(* IEC 61131-3 sources: test/Class/HmiScreen, 1 file *)

(* ---- HmiScreen.st ---- *)
#include "..\..\Source\Common\hmi_nuc.h"

(*!
<Class
	Name               = "HmiScreen"
	Revision           = "0.1"
	RealtimeTask       = "false"
	CyclicTask         = "false"
	BackgroundTask     = "false"
	Sigmatek           = "true"
	OSInterface        = "false"
	HighPriority       = "false"
	Automatic          = "false"
	UpdateMode         = "Prescan"
	SharedCommandTable = "true"
	Objectsize         = "(284,120)">
	<Channels>
		<Client Name="MemCircle" Required="true" Internal="true"/>
		<Client Name="MemImage" Required="true" Internal="true"/>
		<Client Name="MemIO" Required="true" Internal="true"/>
		<Client Name="MemLine" Required="true" Internal="true"/>
		<Client Name="MemRectangle" Required="true" Internal="true"/>
		<Client Name="MemText" Required="true" Internal="true"/>
		<Client Name="MemZorder" Required="true" Internal="true"/>
	</Channels>
	<Dependencies>
		<Files>
			<File Path=".\Source\Common\hmi_nuc.h" Include="true"/>
		</Files>
	</Dependencies>
	<RevDoku>
		<Owner Company="sigmatek" Author="kolott"/>
		<Dokumentation Revision="0.1" Date="2014-04-15" Author="kolott" Company="sigmatek" Description="new method FreeMem()"/>
	</RevDoku>
	<Network Name="HmiScreen">
		<!-- List of Components in this network -->
		<Components>
			<Object
				Name       = "_base"
				Class      = "HmiBaseList"
				Position   = "(218,120)"
				Visualized = "false">
				<Channels>
					<Server Name="ClassSvr"/>
					<Client Name="File"/>
				</Channels>
			</Object>
			<Object
				Name       = "MemCircle"
				Class      = "HmiMemCircle"
				Position   = "(600,510)"
				Visualized = "false">
				<Channels>
					<Server Name="ClassSvr"/>
					<Client Name="File"/>
				</Channels>
			</Object>
			<Object
				Name       = "MemImage"
				Class      = "HmiMemImage"
				Position   = "(600,810)"
				Visualized = "false">
				<Channels>
					<Server Name="ClassSvr"/>
					<Client Name="File"/>
				</Channels>
			</Object>
			<Object
				Name       = "MemIO"
				Class      = "HmiMemIO"
				Position   = "(210,810)"
				Visualized = "false">
				<Channels>
					<Server Name="ClassSvr"/>
					<Client Name="File"/>
				</Channels>
			</Object>
			<Object
				Name       = "MemLine"
				Class      = "HmiMemLine"
				Position   = "(600,660)"
				Visualized = "false">
				<Channels>
					<Server Name="ClassSvr"/>
					<Client Name="File"/>
				</Channels>
			</Object>
			<Object
				Name       = "MemRectangle"
				Class      = "HmiMemRectangle"
				Position   = "(210,510)"
				Visualized = "false">
				<Channels>
					<Server Name="ClassSvr"/>
					<Client Name="File"/>
				</Channels>
			</Object>
			<Object
				Name       = "MemText"
				Class      = "HmiMemText"
				Position   = "(210,660)"
				Visualized = "false">
				<Channels>
					<Server Name="ClassSvr"/>
					<Client Name="File"/>
				</Channels>
			</Object>
			<Object
				Name       = "MemZorder"
				Class      = "HmiMemZorder"
				Position   = "(450,330)"
				Visualized = "false">
				<Channels>
					<Server Name="ClassSvr"/>
					<Client Name="File"/>
				</Channels>
			</Object>
		</Components>
		<Comments>
		</Comments>
		<!-- List of Connections in this network -->
		<Connections>
			<Connection Source="this.ClassSvr" Destination="_base.ClassSvr" Vertices="(1072,210),(518,210),"/>
			<Connection Source="_base.File" Destination="this.File" Vertices="(218,210),(38,210),"/>
			<Connection Source="this.MemZorder" Destination="MemZorder.ClassSvr"/>
			<Connection Source="MemZorder.File" Destination="this.File" Vertices="(450,420),(38,210),"/>
			<Connection Source="this.MemRectangle" Destination="MemRectangle.ClassSvr"/>
			<Connection Source="MemRectangle.File" Destination="this.File" Vertices="(210,600),(38,210),"/>
			<Connection Source="this.MemText" Destination="MemText.ClassSvr"/>
			<Connection Source="MemText.File" Destination="this.File" Vertices="(210,750),(38,210),"/>
			<Connection Source="this.MemIO" Destination="MemIO.ClassSvr"/>
			<Connection Source="MemIO.File" Destination="this.File" Vertices="(210,900),(38,210),"/>
			<Connection Source="this.MemCircle" Destination="MemCircle.ClassSvr"/>
			<Connection Source="MemCircle.File" Destination="this.File" Vertices="(600,600),(38,210),"/>
			<Connection Source="this.MemLine" Destination="MemLine.ClassSvr"/>
			<Connection Source="MemLine.File" Destination="this.File" Vertices="(600,750),(38,210),"/>
			<Connection Source="this.MemImage" Destination="MemImage.ClassSvr"/>
			<Connection Source="MemImage.File" Destination="this.File" Vertices="(600,900),(38,210),"/>
		</Connections>
		<!-- Headerfiles -->
		<Options>
		</Options>
	</Network>
</Class>
*)
#pragma using HmiBaseList

HmiScreen : CLASS
: HmiBaseList
  //Servers:
  //Clients:
	MemRectangle 	: CltChCmd_HmiMemRectangle;
	MemText 	: CltChCmd_HmiMemText;
	MemIO 	: CltChCmd_HmiMemIO;
	MemCircle 	: CltChCmd_HmiMemCircle;
	MemLine 	: CltChCmd_HmiMemLine;
	MemImage 	: CltChCmd_HmiMemImage;
	MemZorder 	: CltChCmd_HmiMemZorder;
  //Variables:
		StartFunct 	: UDINT;
		EndFunct 	: UDINT;
  //Functions:

	FUNCTION VIRTUAL Load
		VAR_OUTPUT
			retcode 	: BOOL;
		END_VAR;

	FUNCTION VIRTUAL Free;

	FUNCTION GLOBAL GetZorder
		VAR_INPUT
			index 	: UDINT;
		END_VAR
		VAR_OUTPUT
			retcode 	: ^HMI_ANYTHING;
		END_VAR;

	FUNCTION GLOBAL GetZorderNo
		VAR_OUTPUT
			retcode 	: UDINT;
		END_VAR;

	FUNCTION GLOBAL GetControl
		VAR_INPUT
			pany 	: ^HMI_ANYTHING;
		END_VAR
		VAR_OUTPUT
			retcode 	: ^void;
		END_VAR;

	FUNCTION GLOBAL GetStartFunct
		VAR_OUTPUT
			retcode 	: UDINT;
		END_VAR;

	FUNCTION GLOBAL GetEndFunct
		VAR_OUTPUT
			retcode 	: UDINT;
		END_VAR;

	FUNCTION GLOBAL FreeMem;
  //Tables:
	FUNCTION @STD
		VAR_OUTPUT
			ret_code	: CONFSTATES;
		END_VAR;
	FUNCTION GLOBAL TAB @CT_;
END_CLASS;

#pragma using HmiMemCircle
#pragma using HmiMemImage
#pragma using HmiMemIO
#pragma using HmiMemLine
#pragma using HmiMemRectangle
#pragma using HmiMemText
#pragma using HmiMemZorder

FUNCTION VIRTUAL HmiScreen::Free

  MemZorder.Free();
  MemRectangle.Free();
  MemText.Free();
  MemIO.Free();
  MemCircle.Free();
  MemLine.Free();
  MemImage.Free();

END_FUNCTION

FUNCTION VIRTUAL HmiScreen::Load
	VAR_OUTPUT
		retcode 	: BOOL;
	END_VAR
  VAR
  	any : HMI_ANYTHING;
    tmp16 : uint;
    room : HMI_ROOM;
  END_VAR

  init_HMI_ANYTHING(#any);
  StartFunct := HMI_DEFSCOPE;
  EndFunct   := HMI_DEFSCOPE;

  File.Read_HMI_ROOM(#room); // position laden

  File.Read_HMI_ANYTHING(#any); // start-funktion laden
  if(any.ima = HMI_IMA_V_FUNCTIONLIST) then
    StartFunct := to_udint(any.value);
  end_if;

  File.Read_HMI_ANYTHING(#any); // ready-funktion laden
  if(any.ima = HMI_IMA_V_FUNCTIONLIST) then
    if(StartFunct = HMI_DEFSCOPE) then
      StartFunct := to_udint(any.value);
    end_if;
  end_if;

  File.Read_HMI_ANYTHING(#any); // run-funktion laden

  File.Read_HMI_ANYTHING(#any); // end-funktion laden
  if(any.ima = HMI_IMA_V_FUNCTIONLIST) then
    EndFunct := to_udint(any.value);
  end_if;

  File.FRead(#tmp16, 2); // firstinput x
  File.FRead(#tmp16, 2); // firstinput y
  File.FRead(#tmp16, 1); // statebits

  MemZorder.Load();
  MemRectangle.Load();
  MemText.Load();
  MemIo.Load();
  MemCircle.Load();
  MemLine.Load();
  MemImage.Load();

//  MemKeypad.Load();

  retcode := File.FChkFile();
  if(retcode = false) then
    Free();
  end_if;

END_FUNCTION

FUNCTION GLOBAL HmiScreen::GetZorder
	VAR_INPUT
		index 	: UDINT;
	END_VAR
	VAR_OUTPUT
		retcode 	: ^HMI_ANYTHING;
	END_VAR

  retcode := MemZorder.Get(index);

END_FUNCTION

FUNCTION GLOBAL HmiScreen::GetZorderNo
	VAR_OUTPUT
		retcode 	: UDINT;
	END_VAR

  retcode := MemZorder.GetNo();

END_FUNCTION

FUNCTION GLOBAL HmiScreen::GetControl
	VAR_INPUT
		pany 	: ^HMI_ANYTHING;
	END_VAR
	VAR_OUTPUT
		retcode 	: ^void;
	END_VAR

  retcode := NIL;
  if(pany <> NIL) then
    case(pany^.ima) of
      HMI_IMA_V_RECTANGLE : retcode := MemRectangle.Get(to_udint(pany^.value));
      HMI_IMA_V_LINE      : retcode := MemLine.Get(to_udint(pany^.value));
      HMI_IMA_V_CIRCLE    : retcode := MemCircle.Get(to_udint(pany^.value));
      HMI_IMA_V_TEXT      : retcode := MemText.Get(to_udint(pany^.value));
      HMI_IMA_V_IMAGE     : retcode := MemImage.Get(to_udint(pany^.value));
      HMI_IMA_V_IO        : retcode := MemIO.Get(to_udint(pany^.value));
    end_case;
  end_if;

END_FUNCTION

FUNCTION GLOBAL HmiScreen::GetStartFunct
	VAR_OUTPUT
		retcode 	: UDINT;
	END_VAR

  retcode := StartFunct;

END_FUNCTION

FUNCTION GLOBAL HmiScreen::GetEndFunct
	VAR_OUTPUT
		retcode 	: UDINT;
	END_VAR

  retcode := EndFunct;

END_FUNCTION

FUNCTION GLOBAL HmiScreen::FreeMem

  Free();

END_FUNCTION
